TYPE "ST_DigitalInputHal"
VERSION : 0.1
   STRUCT
      Value : Bool;
      Quality : Bool := TRUE;
   END_STRUCT;

END_TYPE

